(* IEC 61131-3 sources: plc-cip-batch-control/plc/fb, 6 files *)

(* ---- FB_Alarm.st ---- *)
(*
    FB_Alarm.st: one alarm point, following the ISA-18.2 state model.

    States are held in the ST_Alarm structure the caller owns, so the whole
    alarm list is one array a SCADA client can read in a single request:

        xActive  the process condition is true right now
        xLatched the alarm has been raised and not yet cleared
        xAcked   the operator has acknowledged this occurrence

    An alarm returns to normal only when the condition has gone away *and* it
    has been acknowledged, which is what stops a fleeting condition from
    disappearing off the list before anybody has seen it.
*)

FUNCTION_BLOCK FB_Alarm
VAR_INPUT
    xCondition  : BOOL;
    xEnable     : BOOL := TRUE;
    xAck        : BOOL;
    iPriority   : INT := 3;
    tOnDelay    : TIME := T#0s;
    tOffDelay   : TIME := T#0s;
    rNowS       : REAL;
END_VAR
VAR_IN_OUT
    stAlarm     : ST_Alarm;
END_VAR
VAR_OUTPUT
    xNewAlarm   : BOOL;     (* one scan pulse when it first latches *)
END_VAR
VAR
    fbOn        : TON;
    fbOff       : TOF;
    fbRise      : R_TRIG;
END_VAR

stAlarm.iPriority := iPriority;

fbOn(IN := xCondition AND xEnable, PT := tOnDelay);
fbOff(IN := fbOn.Q, PT := tOffDelay);
stAlarm.xActive := fbOff.Q;

fbRise(CLK := stAlarm.xActive);
xNewAlarm := fbRise.Q;

IF xNewAlarm THEN
    stAlarm.xLatched := TRUE;
    stAlarm.xAcked := FALSE;
    stAlarm.rTimeInS := rNowS;
    stAlarm.iCount := stAlarm.iCount + 1;
END_IF

IF xAck AND stAlarm.xLatched THEN
    stAlarm.xAcked := TRUE;
END_IF

IF stAlarm.xLatched AND NOT stAlarm.xActive AND stAlarm.xAcked THEN
    stAlarm.xLatched := FALSE;
END_IF

END_FUNCTION_BLOCK

(* ---- FB_CipPhase.st ---- *)
(*
    FB_CipPhase.st: the phase engine.

    Every CIP phase is the same four steps with different parameters, so there
    is one engine and the recipe supplies ST_PhaseParams:

        LINEUP     set the valve matrix, prove the circuit is released
        CHARGE     fill the balance tank from the source, dose to strength
        CIRCULATE  hold the wash at temperature and flow, or rinse to a
                   conductivity endpoint
        RECOVER    push the circuit contents back to the source tank or to
                   drain, then stop

    The important idea is in CIRCULATE. The hold timer only advances while
    temperature, flow and concentration are all inside their limits, so ten
    minutes of "hold" means ten minutes of cleaning that actually met the
    specification, not ten minutes on the clock. That accumulated figure is
    what goes in the batch record.
*)

FUNCTION_BLOCK FB_CipPhase
VAR_INPUT
    xExecute    : BOOL;
    xHolding    : BOOL;
    ePhase      : E_Phase;
    stParams    : ST_PhaseParams;
    rTempC      : REAL;     (* return temperature: the coldest point of the circuit *)
    rFlowM3h    : REAL;
    rConcPct    : REAL;
    rDeltaCond  : REAL;     (* return minus supply conductivity, mS/cm *)
    rLevelPct   : REAL;
    xPumpHealthy : BOOL := TRUE;
    rCycleS     : REAL := 0.1;
END_VAR
VAR_OUTPUT
    eStep       : E_PhaseStep;
    stDemand    : ST_Demand;
    xDone       : BOOL;
    xFailed     : BOOL;
    eFail       : E_FailCode;
    rElapsedS   : REAL;
    rHoldAchievedS : REAL;
    stResult    : ST_PhaseResult;
    xInSpec     : BOOL;     (* all cleaning criteria met right now *)
END_VAR
VAR
    fbStart         : R_TRIG;
    fbEndStable     : TON;
    fbFlowLow       : TON;
    fbTempSlow      : TON;
    rStepElapsedS   : REAL;
    rConcSum        : REAL;
    rConcSamples    : REAL;
    rHoldRequiredS  : REAL;
    rMinPhaseS      : REAL;
    rMaxPhaseS      : REAL;
    rRecoverS       : REAL;
    rFillTargetPct  : REAL;
    xSinglePass     : BOOL;
    eActiveReturn   : E_Return;
    xCharged        : BOOL;
    xTempOk         : BOOL;
    xFlowOk         : BOOL;
    xConcOk         : BOOL;
    xDoseDemand     : BOOL;
END_VAR

fbStart(CLK := xExecute);

(* ---- initialise on the rising edge of the execute request ------------- *)
IF fbStart.Q THEN
    eStep := PS_LINEUP;
    rElapsedS := 0.0;
    rStepElapsedS := 0.0;
    rHoldAchievedS := 0.0;
    rConcSum := 0.0;
    rConcSamples := 0.0;
    xCharged := FALSE;
    xDone := FALSE;
    xFailed := FALSE;
    eFail := FC_NONE;
    stResult.ePhase := ePhase;
    stResult.xExecuted := TRUE;
    stResult.xPass := FALSE;
    stResult.eFail := FC_NONE;
    stResult.rDurationS := 0.0;
    stResult.rHoldAchievedS := 0.0;
    stResult.rMinTempC := 999.0;
    stResult.rMaxTempC := -999.0;
    stResult.rMinFlow := 999.0;
    stResult.rMeanConcPct := 0.0;
    stResult.rEndConductivity := 0.0;
    stResult.xAdaptiveEnd := FALSE;
    stResult.rWaterL := 0.0;
    stResult.rChemL := 0.0;
    stResult.rEnergyKWh := 0.0;
END_IF

rHoldRequiredS := TimeToSeconds(stParams.tHold);
rMinPhaseS     := TimeToSeconds(stParams.tMinPhase);
rMaxPhaseS     := TimeToSeconds(stParams.tMaxPhase);
rRecoverS      := TimeToSeconds(stParams.tRecover);

(* An adaptive phase is judged on the conductivity endpoint, so the hold
   requirement does not apply and the record should not imply that it does. *)
stResult.xAdaptiveEnd := stParams.xAdaptiveEnd;
IF stParams.xAdaptiveEnd THEN
    stResult.rHoldRequiredS := 0.0;
ELSE
    stResult.rHoldRequiredS := rHoldRequiredS;
END_IF

(* A recirculating phase makes its charge up in a closed loop through the
   balance tank and only sends the liquid to eReturn when it recovers at the
   end. A single-pass phase runs from the source straight to eReturn, on a
   small working volume so the tank washes out in about a minute. *)
xSinglePass := NOT stParams.xRecirculate;
IF xSinglePass THEN
    rFillTargetPct := C_RINSE_LEVEL_PCT;
ELSE
    rFillTargetPct := C_FILL_TARGET_PCT;
END_IF

IF stParams.xRecirculate AND (eStep <> PS_RECOVER) THEN
    eActiveReturn := RET_BALANCE;
ELSE
    eActiveReturn := stParams.eReturn;
END_IF

(* ---- idle: hold everything closed ------------------------------------ *)
IF NOT xExecute THEN
    stDemand.eSource := SRC_NONE;
    stDemand.eReturn := RET_DRAIN;
    stDemand.rFlowSp := 0.0;
    stDemand.rTempSp := 0.0;
    stDemand.xHeat := FALSE;
    stDemand.xDose := FALSE;
    stDemand.xSupplyPump := FALSE;
    stDemand.xReturnPump := FALSE;
    stDemand.xFillValve := FALSE;
    xInSpec := FALSE;
    RETURN;
END_IF

(* ---- criteria evaluated once, used by several steps ------------------- *)
xTempOk := (NOT stParams.xHeat) OR (rTempC >= stParams.rTempMin);
xFlowOk := rFlowM3h >= stParams.rFlowMin;
xConcOk := (NOT stParams.xDose) OR
           ((rConcPct >= stParams.rConcMin) AND (rConcPct <= stParams.rConcMax));
xInSpec := xTempOk AND xFlowOk AND xConcOk;

(* Dose whenever the strength has drifted below setpoint. Above the band the
   valve simply stays shut; the phase dilutes back with the next charge. *)
xDoseDemand := stParams.xDose AND (rConcPct < stParams.rConcSp);

(* ---- the line-up is common to every running step ---------------------- *)
stDemand.eSource := stParams.eSource;
stDemand.eReturn := eActiveReturn;
stDemand.rTempSp := stParams.rTempSp;
stDemand.rFlowSp := stParams.rFlowSp;

IF xHolding THEN
    (* Freeze: keep the valve matrix so the circuit stays full but stop
       circulating, stop heating and stop dosing. Accumulators do not advance,
       so a held phase does not earn hold time. *)
    stDemand.xSupplyPump := FALSE;
    stDemand.xReturnPump := TRUE;
    stDemand.xHeat := FALSE;
    stDemand.xDose := FALSE;
    stDemand.xFillValve := FALSE;
    RETURN;
END_IF

rElapsedS := rElapsedS + rCycleS;
rStepElapsedS := rStepElapsedS + rCycleS;
stResult.rDurationS := rElapsedS;

(* ---- the step machine ------------------------------------------------- *)
CASE eStep OF

    PS_LINEUP:
        stDemand.xSupplyPump := FALSE;
        stDemand.xReturnPump := TRUE;
        stDemand.xHeat := FALSE;
        stDemand.xDose := FALSE;
        stDemand.xFillValve := TRUE;
        IF rStepElapsedS >= 5.0 THEN
            eStep := PS_CHARGE;
            rStepElapsedS := 0.0;
        ELSIF rStepElapsedS > 60.0 THEN
            eFail := FC_LINEUP_TIMEOUT;
        END_IF

    PS_CHARGE:
        stDemand.xReturnPump := TRUE;
        stDemand.xFillValve := rLevelPct < rFillTargetPct;
        (* Start circulating as soon as there is enough suction head; the
           remaining fill and the dose trim happen while the pump runs, which
           is also what satisfies the no-dosing-without-flow interlock. *)
        stDemand.xSupplyPump := rLevelPct >= C_PUMP_START_PCT;
        stDemand.xHeat := stParams.xHeat AND stDemand.xSupplyPump;
        stDemand.xDose := xDoseDemand AND stDemand.xSupplyPump;
        xCharged := (rLevelPct >= rFillTargetPct) AND xConcOk;
        IF xCharged THEN
            eStep := PS_CIRCULATE;
            rStepElapsedS := 0.0;
        ELSIF rStepElapsedS > 600.0 THEN
            eFail := FC_CHARGE_TIMEOUT;
        END_IF

    PS_CIRCULATE:
        stDemand.xSupplyPump := TRUE;
        stDemand.xReturnPump := TRUE;
        stDemand.xHeat := stParams.xHeat;
        stDemand.xDose := xDoseDemand;
        (* Single-pass phases keep drawing fresh liquid; recirculating phases
           only top up if the circuit has swallowed some of the charge. *)
        stDemand.xFillValve := rLevelPct < rFillTargetPct;

        IF xInSpec THEN
            rHoldAchievedS := rHoldAchievedS + rCycleS;
        END_IF
        stResult.rHoldAchievedS := rHoldAchievedS;

        (* Statistics start once the loop has settled, otherwise every phase
           records the pump ramp as its minimum flow. *)
        IF rStepElapsedS > 15.0 THEN
            IF rTempC < stResult.rMinTempC THEN
                stResult.rMinTempC := rTempC;
            END_IF
            IF rTempC > stResult.rMaxTempC THEN
                stResult.rMaxTempC := rTempC;
            END_IF
            IF rFlowM3h < stResult.rMinFlow THEN
                stResult.rMinFlow := rFlowM3h;
            END_IF
            rConcSum := rConcSum + rConcPct;
            rConcSamples := rConcSamples + 1.0;
            stResult.rMeanConcPct := rConcSum / rConcSamples;
        END_IF
        stResult.rEndConductivity := rDeltaCond;

        (* Endpoint. An adaptive rinse stops when the return water is as clean
           as the water going in; everything else stops on verified hold time. *)
        fbEndStable(IN := stParams.xAdaptiveEnd AND (rDeltaCond <= stParams.rEndConductivity)
                          AND (rElapsedS >= rMinPhaseS),
                    PT := T#10s);

        IF stParams.xAdaptiveEnd THEN
            IF fbEndStable.Q THEN
                eStep := PS_RECOVER;
                rStepElapsedS := 0.0;
            ELSIF rElapsedS >= rMaxPhaseS THEN
                eFail := FC_RINSE_NOT_CLEAN;
            END_IF
        ELSE
            IF rHoldAchievedS >= rHoldRequiredS THEN
                eStep := PS_RECOVER;
                rStepElapsedS := 0.0;
            ELSIF rElapsedS >= rMaxPhaseS THEN
                eFail := FC_PHASE_TIMEOUT;
            END_IF
        END_IF

        (* Sustained excursions are faults, not just missing hold time. *)
        fbFlowLow(IN := NOT xFlowOk, PT := T#60s);
        IF fbFlowLow.Q THEN
            eFail := FC_FLOW_LOW;
        END_IF
        fbTempSlow(IN := stParams.xHeat AND NOT xTempOk, PT := T#8m);
        IF fbTempSlow.Q THEN
            eFail := FC_TEMP_TIMEOUT;
        END_IF
        IF rLevelPct < C_LEVEL_TRIP_PCT THEN
            eFail := FC_LEVEL_LOW;
        END_IF

    PS_RECOVER:
        (* Push the contents back where they came from. Heat and dose are off
           and the fill valve is shut, so the balance tank drains as the pump
           empties it into the return line. Draining it properly is what keeps
           the next phase's charge from being diluted by the last one's
           chemical and what keeps the following rinse short. *)
        stDemand.xSupplyPump := (rStepElapsedS < rRecoverS)
                                AND (rLevelPct > C_PUMP_START_PCT);
        stDemand.xReturnPump := TRUE;
        stDemand.xHeat := FALSE;
        stDemand.xDose := FALSE;
        stDemand.xFillValve := FALSE;
        IF (rStepElapsedS >= rRecoverS) OR (rLevelPct <= C_PUMP_START_PCT) THEN
            eStep := PS_DONE;
            rStepElapsedS := 0.0;
        END_IF

    PS_DONE:
        stDemand.xSupplyPump := FALSE;
        stDemand.xReturnPump := FALSE;
        stDemand.xHeat := FALSE;
        stDemand.xDose := FALSE;
        stDemand.xFillValve := FALSE;
        stDemand.eSource := SRC_NONE;
        xDone := TRUE;
        stResult.xPass := TRUE;
END_CASE

IF NOT xPumpHealthy THEN
    eFail := FC_PUMP_FAULT;
END_IF

IF eFail <> FC_NONE THEN
    xFailed := TRUE;
    xDone := FALSE;
    eStep := PS_DONE;
    stResult.xPass := FALSE;
    stResult.eFail := eFail;
    stDemand.xSupplyPump := FALSE;
    stDemand.xReturnPump := FALSE;
    stDemand.xHeat := FALSE;
    stDemand.xDose := FALSE;
    stDemand.xFillValve := FALSE;
END_IF

END_FUNCTION_BLOCK

(* ---- FB_Pid.st ---- *)
(*
    FB_Pid.st: PI(D) controller with clamping anti-windup.

    The integral only accumulates while the output is off its limit, which is
    what keeps the steam valve from winding up during the long fill step and
    then overshooting the wash temperature when circulation finally starts.

    rTi and rTd are in seconds. rTi = 0 disables the integral term.
*)

FUNCTION_BLOCK FB_Pid
VAR_INPUT
    xEnable     : BOOL;
    rPv         : REAL;
    rSp         : REAL;
    rKp         : REAL := 1.0;
    rTi         : REAL := 0.0;
    rTd         : REAL := 0.0;
    rOutMin     : REAL := 0.0;
    rOutMax     : REAL := 100.0;
    rCycleS     : REAL := 0.1;
END_VAR
VAR_OUTPUT
    rOut        : REAL;
    rError      : REAL;
    xSaturated  : BOOL;
END_VAR
VAR
    rIntegral   : REAL;
    rPrevPv     : REAL;
    xFirstScan  : BOOL := TRUE;
    rDerivative : REAL;
    rRaw        : REAL;
END_VAR

IF NOT xEnable THEN
    (* Bumpless enough for this duty: park the integrator and the output. *)
    rIntegral := 0.0;
    rOut := rOutMin;
    rError := 0.0;
    xSaturated := FALSE;
    xFirstScan := TRUE;
    rPrevPv := rPv;
    RETURN;
END_IF

rError := rSp - rPv;

(* Derivative on the measurement, so a setpoint step does not kick the valve. *)
IF xFirstScan THEN
    rDerivative := 0.0;
    xFirstScan := FALSE;
ELSIF rCycleS > 0.0 THEN
    rDerivative := (rPrevPv - rPv) / rCycleS;
ELSE
    rDerivative := 0.0;
END_IF
rPrevPv := rPv;

rRaw := rKp * rError + rIntegral + rKp * rTd * rDerivative;

(* Clamping anti-windup: integrate only if that does not push further into a
   limit the output is already sitting on. *)
IF rTi > 0.0 THEN
    IF (rRaw < rOutMax) AND (rRaw > rOutMin) THEN
        rIntegral := rIntegral + (rKp / rTi) * rError * rCycleS;
    ELSIF (rRaw >= rOutMax) AND (rError < 0.0) THEN
        rIntegral := rIntegral + (rKp / rTi) * rError * rCycleS;
    ELSIF (rRaw <= rOutMin) AND (rError > 0.0) THEN
        rIntegral := rIntegral + (rKp / rTi) * rError * rCycleS;
    END_IF
    rIntegral := LIMIT(rOutMin - rOutMax, rIntegral, rOutMax - rOutMin);
END_IF

rRaw := rKp * rError + rIntegral + rKp * rTd * rDerivative;
rOut := LIMIT(rOutMin, rRaw, rOutMax);
xSaturated := (rRaw > rOutMax) OR (rRaw < rOutMin);

END_FUNCTION_BLOCK

(* ---- FB_Pump.st ---- *)
(*
    FB_Pump.st: motor starter with interlock, feedback supervision and a
    latched trip.

    A pump that is commanded to run but reports no feedback inside
    tFeedbackTimeout latches a trip. Clearing it needs an explicit reset, not
    just the disappearance of the fault, so an intermittent contactor cannot
    silently restart the skid mid-wash.
*)

FUNCTION_BLOCK FB_Pump
VAR_INPUT
    xStart              : BOOL;
    xInterlockOk        : BOOL;
    xRunFeedback        : BOOL;
    xFault              : BOOL;     (* motor protection relay *)
    xReset              : BOOL;
    tFeedbackTimeout    : TIME := T#5s;
END_VAR
VAR_OUTPUT
    xRun                : BOOL;     (* to the field *)
    xTripped            : BOOL;
    xFeedbackFault      : BOOL;
    xHealthy            : BOOL;
END_VAR
VAR
    fbFeedback  : TON;
    fbFault     : R_TRIG;
END_VAR

fbFault(CLK := xFault);

IF fbFault.Q THEN
    xTripped := TRUE;
END_IF

IF xReset AND NOT xFault THEN
    xTripped := FALSE;
    xFeedbackFault := FALSE;
END_IF

xRun := xStart AND xInterlockOk AND NOT xTripped AND NOT xFeedbackFault;

(* Supervise only the commanded direction: a pump that keeps running after the
   command drops is a separate condition, alarmed in PRG_Alarms. *)
fbFeedback(IN := xRun AND NOT xRunFeedback, PT := tFeedbackTimeout);
IF fbFeedback.Q THEN
    xFeedbackFault := TRUE;
    xRun := FALSE;
END_IF

xHealthy := NOT xTripped AND NOT xFeedbackFault AND NOT xFault;

END_FUNCTION_BLOCK

(* ---- FB_Totaliser.st ---- *)
(*
    FB_Totaliser.st: rectangular integration of a rate against the scan
    period, with a low-flow cut-off.

    The cut-off matters: a flow transmitter parked at 0.3 m3/h of noise while
    the pump is stopped would otherwise book about 7 litres an hour of water
    that never moved and those litres end up in the batch record.
*)

FUNCTION_BLOCK FB_Totaliser
VAR_INPUT
    xEnable     : BOOL;
    rRatePerHour : REAL;
    rCutOff     : REAL := 0.0;
    rCycleS     : REAL := 0.1;
    xReset      : BOOL;
END_VAR
VAR_OUTPUT
    rTotal      : REAL;
    rRateUsed   : REAL;
END_VAR

IF xReset THEN
    rTotal := 0.0;
END_IF

IF xEnable AND (rRatePerHour > rCutOff) THEN
    rRateUsed := rRatePerHour;
    rTotal := rTotal + rRatePerHour * rCycleS / 3600.0;
ELSE
    rRateUsed := 0.0;
END_IF

END_FUNCTION_BLOCK

(* ---- FB_UnitStateMachine.st ---- *)
(*
    FB_UnitStateMachine.st: the ISA-88 unit procedural state model.

    Commands are edge triggered, so a stuck HMI bit cannot hold the unit in a
    transition. ABORTING is deliberately not instantaneous: it runs for
    tAbortSettle so the control layer can shut the steam valve and stop the
    pumps in a defined order before the unit is declared ABORTED.

        IDLE -> STARTING -> RUNNING -> COMPLETING -> COMPLETE -> IDLE
                              |  ^
                          HOLDING |
                              |  RESTARTING
                              v  |
                            HELD +
        any active state -> ABORTING -> ABORTED -> IDLE
*)

FUNCTION_BLOCK FB_UnitStateMachine
VAR_INPUT
    xStart              : BOOL;
    xHold               : BOOL;
    xRestart            : BOOL;
    xAbort              : BOOL;
    xReset              : BOOL;
    xReadyToStart       : BOOL;
    xProcedureComplete  : BOOL;
    xProcedureFailed    : BOOL;
    xSafetyTrip         : BOOL;
    tAbortSettle        : TIME := T#5s;
    tHoldSettle         : TIME := T#2s;
END_VAR
VAR_OUTPUT
    eState              : E_UnitState;
    xExecute            : BOOL;     (* the phase engine may run *)
    xHolding            : BOOL;     (* freeze the phase, keep the line-up *)
    xAborting           : BOOL;
    xStartPulse         : BOOL;     (* one scan, initialise the procedure *)
    xActive             : BOOL;     (* anything other than IDLE/COMPLETE/ABORTED *)
END_VAR
VAR
    fbStart     : R_TRIG;
    fbHold      : R_TRIG;
    fbRestart   : R_TRIG;
    fbAbort     : R_TRIG;
    fbReset     : R_TRIG;
    fbAbortTmr  : TON;
    fbHoldTmr   : TON;
END_VAR

fbStart(CLK := xStart);
fbHold(CLK := xHold);
fbRestart(CLK := xRestart);
fbAbort(CLK := xAbort);
fbReset(CLK := xReset);

xStartPulse := FALSE;

(* An abort request or a safety trip pre-empts every other transition. *)
IF (fbAbort.Q OR xSafetyTrip OR xProcedureFailed)
   AND (eState <> UST_IDLE) AND (eState <> UST_COMPLETE)
   AND (eState <> UST_ABORTED) AND (eState <> UST_ABORTING) THEN
    eState := UST_ABORTING;
END_IF

CASE eState OF
    UST_IDLE:
        (* Park both settle timers so a previous batch cannot leave one
           already elapsed and collapse the next HOLDING into one scan. *)
        fbHoldTmr(IN := FALSE, PT := tHoldSettle);
        fbAbortTmr(IN := FALSE, PT := tAbortSettle);
        IF fbStart.Q AND xReadyToStart THEN
            eState := UST_STARTING;
        END_IF

    UST_STARTING:
        xStartPulse := TRUE;
        eState := UST_RUNNING;

    UST_RUNNING:
        IF xProcedureComplete THEN
            eState := UST_COMPLETING;
        ELSIF fbHold.Q THEN
            eState := UST_HOLDING;
        END_IF

    UST_HOLDING:
        fbHoldTmr(IN := TRUE, PT := tHoldSettle);
        IF fbHoldTmr.Q THEN
            fbHoldTmr(IN := FALSE, PT := tHoldSettle);
            eState := UST_HELD;
        END_IF

    UST_HELD:
        IF fbRestart.Q THEN
            eState := UST_RESTARTING;
        END_IF

    UST_RESTARTING:
        eState := UST_RUNNING;

    UST_COMPLETING:
        eState := UST_COMPLETE;

    UST_COMPLETE:
        IF fbReset.Q THEN
            eState := UST_IDLE;
        END_IF

    UST_ABORTING:
        fbAbortTmr(IN := TRUE, PT := tAbortSettle);
        IF fbAbortTmr.Q THEN
            fbAbortTmr(IN := FALSE, PT := tAbortSettle);
            eState := UST_ABORTED;
        END_IF

    UST_ABORTED:
        IF fbReset.Q AND NOT xSafetyTrip THEN
            eState := UST_IDLE;
        END_IF
END_CASE

xExecute  := (eState = UST_RUNNING);
(* RESTARTING counts as holding. It lasts one scan, and the phase has not
   resumed yet, so the phase engine must keep its state through it. Leaving it
   out of both outputs gives the engine one scan in which it is neither
   executing nor holding, which it reads as the phase having ended; the next
   scan then looks like a fresh start and the phase begins again from zero. *)
xHolding  := (eState = UST_HOLDING) OR (eState = UST_HELD) OR (eState = UST_RESTARTING);
xAborting := (eState = UST_ABORTING);
xActive   := (eState <> UST_IDLE) AND (eState <> UST_COMPLETE) AND (eState <> UST_ABORTED);

END_FUNCTION_BLOCK
